RoboDK station: hand_motion.rdk

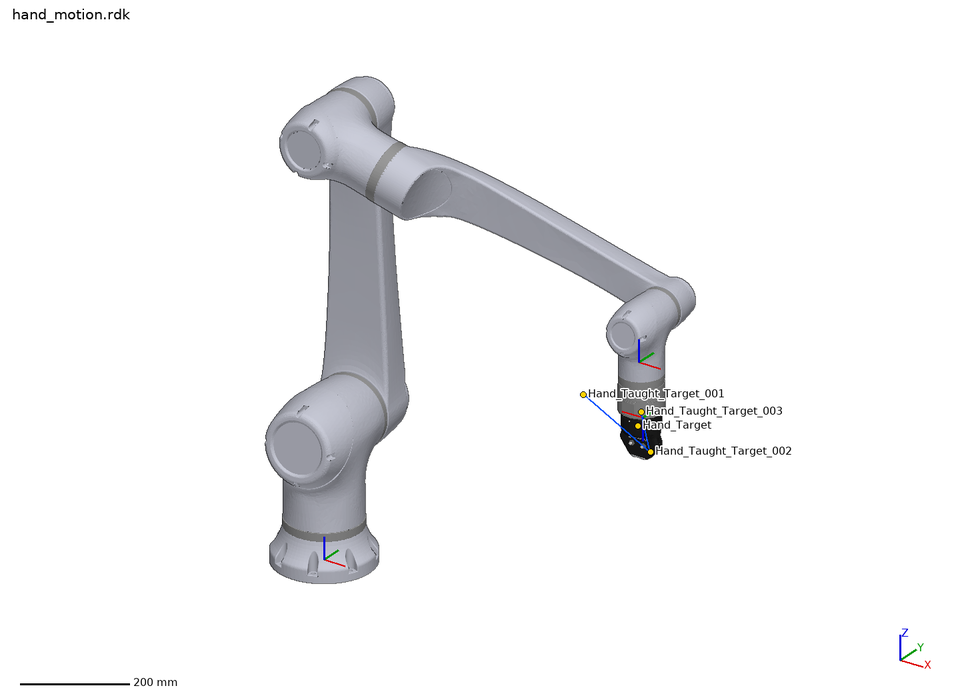
[picture v0: the station drawn from its stored meshes, robots at their saved joint values, targets as dots, program paths as lines]
Station hand_motion (saved by RoboDK 6.0.6). Poses are relative to the parent item; angles as X-Y-Z fixed-axis rotations.
  - frame Neura LARA 8 Base at (0, 0, 0) mm
    - robot Neura LARA 8: 6 axes
        modified DH rows (alpha deg, a mm, theta deg, d mm): 0, 0, 0, 260; -90, 0, -90, 0; 0, 600, -90, 0; -90, 0, 0, 700; 90, 0, 0, 0; -90, 0, 180, 179.5
        joint limits [-180, -135, -155, -180, -180, -360] to [180, 135, 155, 180, 180, 360]; home [0, 0, 90, 0, 90, 0]; saved at [4.66, 0.284, 107.692, 0, 72.024, 4.66]
      - robot RobotiQ 2F-85 Gripper (Mechanism) (model RobotiQ 2F85): 1 axes, payload 5 kg
          joint limits [0] to [85]; home [85]; saved at [0]
        - frame Grip_Attach_Frame at (-4.53, -1.14, 10.96) mm
    - target Hand_Target (Cartesian target) at (661.09, 52.97, 434.07) mm, rotated rx 180 ry 0 rz -180 deg; joints [-5.022, -5.904, 101.187, 0, 84.717, -5.022] of Neura LARA 8
    - target Hand_Taught_Target_001 (Cartesian target) at (618.83, -60.29, 531.83) mm, rotated rx 180 ry 0 rz -180 deg; joints [-5.564, -6.026, 108.01, 0, 78.016, -5.564] of Neura LARA 8
    - target Hand_Taught_Target_002 (Cartesian target) at (718.54, 10.09, 414.63) mm, rotated rx 180 ry 0 rz -180 deg; joints [0.805, 6.645, 105.321, 0, 68.034, 0.805] of Neura LARA 8
    - target Hand_Taught_Target_003 (Cartesian target) at (666.6, 54.33, 464.46) mm, rotated rx 180 ry 0 rz -180 deg; joints [4.66, 0.284, 107.692, 0, 72.024, 4.66] of Neura LARA 8
  - object Cube 50mm at (805.02, 3.79, 48.01) mm, rotated rx 180 ry 0 rz -174.82 deg, size 50 x 50 x 50 mm, geometry from Cube-50mm.sld
  - frame RobotiQ 2F-85 Gripper (Mechanism) Base at (0, 1000, 0) mm
  - program Hand_Taught_Program_172056 (3 instructions, listed below)
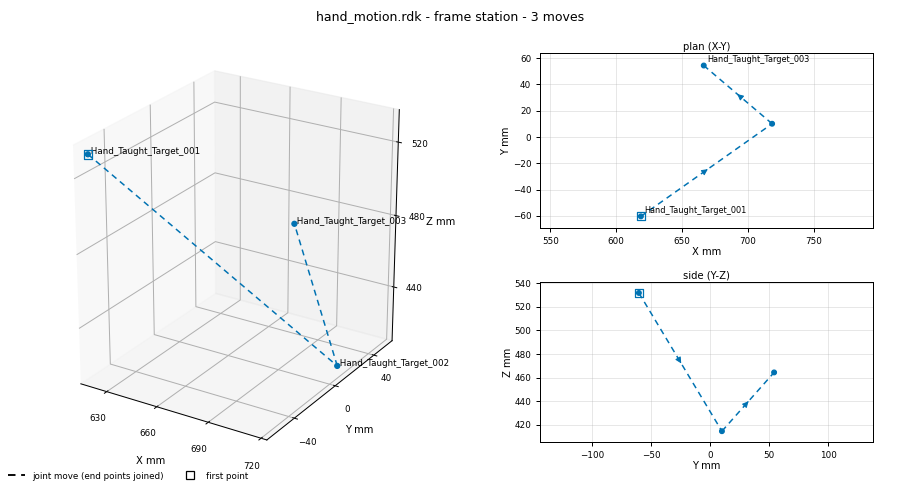
[picture p0: tool path of hand_motion.rdk in frame station, 3 of 3 moves have a stored position in this frame; points joined in program order, loops and branches not executed]

--- program Hand_Taught_Program_172056 (robot Neura LARA 8) ---
  MoveJ (Hand_Taught_Target_001)
  MoveJ (Hand_Taught_Target_002)
  MoveJ (Hand_Taught_Target_003)
